(* IEC 61131-3 sources: LASAL/Class/_DriveMngBase (part 2) *)

           ret_code := READY;

           // Daten werden gelöscht :
           L2Buffer[IntRdIndex].AxisNo := 0;
           L2Buffer[IntRdIndex].bActive := FALSE;
           L2NewEntry -= 1;
           if L2NewEntry < 0 then
            L2NewEntry := 0;
           end_if;
           exit;
        end_if;
      end_for;

    end_if;

  else
    ret_code := NewInst(pPara, pResult);
  end_case;

END_FUNCTION

FUNCTION GLOBAL _DriveMngBase::GetAxisWrPtr
	VAR_INPUT
		usAxis 	: USINT;
	END_VAR
	VAR_OUTPUT
		ptr 	: ^_VaranDriveBase::t_WriteValuePtr;
	END_VAR
  VAR
    MyPara   : CmdStruct;
    MyResult : results;
  END_VAR

  if usAxis >= 0 & usAxis < SDDMAXENTRIES then //HasHan
    if bVaranConnected then
      ptr := toVaran.GetAxisWrPtr(AxisNr:=AxBuffer[usAxis].AxisIndex);
    else
      MyPara.uiCmd    := BUSIF_DRIVEMNGBASE_GET_AXIS_WR_PTR;
      MyPara.aPara[0] := to_dint(AxBuffer[usAxis].AxisIndex);
      ToBusIF.NewInst(#MyPara, #MyResult);
      ptr := MyResult.aData[0]$^_VaranDriveBase::t_WriteValuePtr;
    end_if;
  end_if;

END_FUNCTION

FUNCTION GLOBAL _DriveMngBase::GetAxisRdPtr
	VAR_INPUT
		usAxis 	: USINT;
	END_VAR
	VAR_OUTPUT
		ptr 	: ^_VaranDriveBase::t_ReadValuePtr;
	END_VAR
  VAR
    MyPara   : CmdStruct;
    MyResult : results;
  END_VAR

  if usAxis >= 0 & usAxis < SDDMAXENTRIES then //HasHan
    if bVaranConnected then
      ptr := toVaran.GetAxisRdPtr(AxisNr:=AxBuffer[usAxis].AxisIndex);
    else
      MyPara.uiCmd    := BUSIF_DRIVEMNGBASE_GET_AXIS_RD_PTR;
      MyPara.aPara[0] := to_dint(AxBuffer[usAxis].AxisIndex);
      ToBusIF.NewInst(#MyPara, #MyResult);
      ptr := MyResult.aData[0]$^_VaranDriveBase::t_ReadValuePtr;
    end_if;
  end_if;

END_FUNCTION

FUNCTION GLOBAL _DriveMngBase::InitDrive
	VAR_INPUT
		Mode 	: USINT;
	END_VAR
  VAR
    UserPara     : CmdStruct;
    UserResult   : Results;
    x            : USINT;
    pThisNewInst : ^void;
  END_VAR

  if bVaranConnected then
    toVaran.InitDrive();
  else
    UserPara.uiCmd := BUSIF_DRIVEMNGBASE_INIT_DRIVE;
    ToBusIF.NewInst(#UserPara, #UserResult);
  end_if;

  for x := 0 to (SDDMAXENTRIES - 1) do
    if (AxBuffer[x].pThis <> NIL) then
      if (AxBuffer[x].AxisOk = 1) then
        if Mode = 0 then
          UserPara.uiCmd := SDD_INITAXLE;
        else
          UserPara.uiCmd := SDD_URINITAXLE;
        end_if;

        pThisNewInst := AxBuffer[x].pThis;
        pThisNewInst$^VirtualBase^.NewInst(#UserPara, #UserResult);
      end_if;
    end_if;
  end_for;

END_FUNCTION

FUNCTION _DriveMngBase::GetAxIndex
	VAR_INPUT
		AxisNo 	: USINT;
	END_VAR
	VAR_OUTPUT
		AxIndex 	: USINT;
	END_VAR
  VAR
  	x     : USINT;
  END_VAR

  AxIndex := 16#FF;

  for x := 0 to (SDDMAXENTRIES - 1) do
    if (AxBuffer[x].pThis <> NIL) then
      if (AxBuffer[x].AxisOk = 1) & (AxBuffer[x].AxisIndex = AxisNo) then
        AxIndex := x;
        exit;
      end_if;
    else
      exit;
    end_if;
  end_for;

END_FUNCTION

FUNCTION _DriveMngBase::GetAxIndexByAxisBit
	VAR_INPUT
		AxisBit 	: BDINT;
	END_VAR
	VAR_OUTPUT
		AxIndex 	: USINT;
	END_VAR
  VAR
  	x     : USINT;
  END_VAR

  AxIndex := 16#FF;

  for x := 0 to (SDDMAXENTRIES - 1) do
    if (AxBuffer[x].pThis <> NIL) then
      if (AxBuffer[x].AxisBit = AxisBit) then
        AxIndex := x;
        exit;
      end_if;
    else
      exit;
    end_if;
  end_for;

END_FUNCTION

FUNCTION _DriveMngBase::GetFirstAxIndex
	VAR_OUTPUT
		AxIndex 	: USINT;
	END_VAR
  VAR
  	x     : USINT;
  END_VAR

  AxIndex := 16#FF;

  for x := 0 to (SDDMAXENTRIES - 1) do
    if (AxBuffer[x].pThis <> NIL) then
      if (AxBuffer[x].AxisOk = 1) then
        AxIndex := x;
        exit;
      end_if;
    else
      exit;
    end_if;
  end_for;

END_FUNCTION

FUNCTION _DriveMngBase::SetFwVersion
VAR
	szValue     : ARRAY[0..19] of CHAR;
  StrLen      : UDINT;
END_VAR

  Bin2Ascii(pt:=#szValue[0], value:=FwVersionInt, format:=16#820);
  StrLen := _strlen(#szValue[0]);
  FwNumStr.WriteDataOff(udLen:= Strlen, udOff:=0, pData:= #szValue[0]);

END_FUNCTION

FUNCTION _DriveMngBase::SetFwDate
VAR
	szValue     : ARRAY[0..19] of CHAR;
  szFwDate    : ARRAY[0..99] of CHAR;
  StrLen      : UDINT;
  Value       : UDINT;
  tmpYear     : UDINT;
END_VAR

  // Ermitteln des Tages
  Value := FWDateInt AND 16#003F0000;
  Value := Value SHR 16;
  Bin2Ascii(pt:=#szValue[0], value:=Value$DINT, format:=16#102);
  _strcpy(#szFwDate[0], #szValue[0]);
  _strcat(#szFwDate[0], ".");

  // ermitteln des Monats
  Value := FWDateInt AND 16#0F000000;
  Value := Value SHR 24;
  Bin2Ascii(pt:=#szValue[0], value:=Value$DINT, format:=16#102);
  _strcat(#szFwDate[0], #szValue[0]);
  _strcat(#szFwDate[0], ".");

  // ermitteln des Jahres
  Value := FWDateInt AND 16#F0000000;
  Value := Value SHR 28;

  //Newer firmwares >= 2016 are using 2 Bits more, which where originally reserved for day, to have more bits to display year dates.
  //With this change we can display year dates until 2063 instead of 2015,
  tmpYear := FWDateInt AND 16#00C00000;
  tmpYear := tmpYear SHR 18; //Shift Right 18 instead of 22 because these two bits are bit 4 and 5 for the year
  Value := Value OR tmpYear;

  Value += 2000;
  Bin2Ascii(pt:=#szValue[0], value:=Value$DINT, format:=16#800);
  _strcat(#szFwDate[0], #szValue[0]);
  _strcat(#szFwDate[0], " ");

  // ermitteln der Stunde
  Value := FWDateInt AND 16#0000FF00;
  Value := Value SHR 8;
  Bin2Ascii(pt:=#szValue[0], value:=Value$DINT, format:=16#102);
  _strcat(#szFwDate[0], #szValue[0]);
  _strcat(#szFwDate[0], ":");

  // ermitteln der Minuten
  Value := FWDateInt AND 16#000000FF;
  Bin2Ascii(pt:=#szValue[0], value:=Value$DINT, format:=16#102);
  _strcat(#szFwDate[0], #szValue[0]);

  StrLen := _strlen(#szFwDate[0]);
  FwDatetr.WriteDataOff(udLen:= Strlen, udOff:=0, pData:= #szFwDate[0]);

END_FUNCTION

(*
Der String kann folgendermaßen formatiert werden.
xxxx 0000 0000 0000     xxxx = keine Funktion.
     .... .... ****     Anzahl der Dezimalstellen.
     .... **** ....     Position des Dezimalpunkts.
     ...* .... ....     Vornullen (Anzahl der Dezimalstellen).
     ..*. .... ....     Nachkomma Nullen.
     .*.. .... ....     Vorzeichen unmittelbar vor wert (-3 ansonsten - 3).
     *... .... ....     Anzahl der Stellen automatisch ermitteln.

*)

FUNCTION _DriveMngBase::Bin2Ascii
	VAR_INPUT
		pt 	: ^CHAR;
		value 	: DINT;
		format 	: BINT;
	END_VAR
VAR
	tmp		: DINT;
	nk		: UINT;
	dig		: UINT;
	hp     : ^CHAR;
	pd     : UINT;
	h      : UINT;
END_VAR

	if((format AND 16#000F) = 0) then
		format := format OR 16#0800;
	end_if;

	if(format AND 16#0800) then
		tmp  := value;
		if tmp = 0 then
			dig := 1;
		else
			dig := 0;
		end_if;

	    while(tmp) do

			tmp := tmp / 10;
			dig += 1;
	    end_while;

	    nk := ((format SHR 4) AND 16#0F);

		if(nk >= dig) then
	      dig := nk + 1;
		end_if;

		format := (format AND 16#FFF0) OR (dig AND 16#000F);
	end_if;

  dig := (format and 16#0F);		// Anzahl der Stellen
  hp  := pt + dig; 					// pointer auf String-Ende
  tmp := value; 					// Zahl
  pd  := (format shr 4) and 16#0F;	// position des Komma

  if(value < 0) then  		// kontrolle ob Zahl negativ
	hp    += 1;
    value := -value;		// Zahl * (-1)
    pt^   := '-';			// Erstes Zeichen auf '-' setzen
  end_if;

  if(format and 16#0200) then   // Nachnullen löschen
    h := pd;
	while(h) do					// Nur Nullen hinter Komma
	  h -= 1;
	  if((value mod 10) = 0) then	// Ist Ziffer Null?
	    value := value / 10; 	// wenn ja, Null löschen
		pd -= 1;
      else
	    h := 0;
      end_if;

	end_while;
  end_if;

  if(pd <> 0) then    	// Komma noch zu setzen?
    hp += 1;
  end_if;

  hp^ := 0;           	// String mit Ascii-0 abschließen
  hp  -= 1;

  repeat
    hp^   := '0' + TO_USINT(value mod 10); //akt. Ziffer
	hp    -= 1;
	pd    -= 1;
	dig   -= 1;
	if(pd = 0)then		//	Komma setzen?
	  hp^ := '.';
	  hp -= 1;
    end_if;

    value := value / 10; 	// nächste Ziffer

    if((dig = 0) & (value <> 0)) then	// Zahl zu groß
	  pt^   := '?'; 	// Formatfehler
	  value := 0;
	end_if;
  until(value = 0) end_repeat;

  if(dig > 0) then 	// mit Vornullen auffüllen
	repeat			// so lange bis Digits auf Null
      if((format and 16#0100)|(pd$INT >= 0)) then   // Vornullen im
        hp^ := '0'; 								// Format angegeben?
      else			// formatfehler (digit zu groß und keine Vornullen)
	    pt^   := '?'; 	// Formatfehler
	    value := 0;
      end_if;
      pd -= 1;
	  hp -= 1;
      if(pd = 0) then	// Komma setzen
	    hp^ := '.';
	    hp -= 1;
      end_if;
	  dig -= 1;
	until(dig = 0) end_repeat; 	// letzte Ziffer?
  end_if;

END_FUNCTION

FUNCTION VIRTUAL GLOBAL _DriveMngBase::RetryCounter::Read
	VAR_OUTPUT
		output (EAX) 	: UDINT;
	END_VAR
  VAR
    MyPara   : CmdStruct;
    MyResult : results;
  END_VAR

  if bVaranConnected then
    RetryCounter := toVaran.RetryCounter.Read();
  else
    MyPara.uiCmd  := BUSIF_DRIVEMNGBASE_READ_RETRY_COUNTER;
    ToBusIF.NewInst(#MyPara, #MyResult);
    RetryCounter := MyResult.aData[0]$UDINT;
  end_if;

  output := RetryCounter;

END_FUNCTION

FUNCTION GLOBAL _DriveMngBase::SetSyncEntry
	VAR_INPUT
		usAxis 	: USINT;
		usValue 	: USINT;
		usPData 	: DINT;
	END_VAR
	VAR_OUTPUT
		retcode 	: DINT;
	END_VAR
  VAR
    MyPara   : CmdStruct;
    MyResult : results;
  END_VAR

  if usAxis >= 0 & usAxis < SDDMAXENTRIES then //HasHan
    if bVaranConnected then
      retcode:=toVaran.SetSyncParameter(us_Axis:=AxBuffer[usAxis].AxisIndex, us_value:=usValue, sd_data:=usPData);
    else
      MyPara.uiCmd    := BUSIF_DRIVEMNGBASE_SET_SYNC_PARA;
      MyPara.aPara[0] := to_dint(AxBuffer[usAxis].AxisIndex);
      MyPara.aPara[1] := to_dint(usValue);
      MyPara.aPara[2] := to_dint(usPData);

      ToBusIF.NewInst(#MyPara, #MyResult);
      retcode := MyResult.aData[0]$DINT;
    end_if;
  else
    retcode := -1;
  end_if;

END_FUNCTION

FUNCTION GLOBAL _DriveMngBase::GetSyncEntry
	VAR_INPUT
		usAxis 	: USINT;
		usValue : USINT;
		usPData : ^DINT;
	END_VAR
	VAR_OUTPUT
		retcode : DINT;
	END_VAR
  VAR
    MyPara   : CmdStruct;
    MyResult : results;
  END_VAR

  if usAxis >= 0 & usAxis < SDDMAXENTRIES then //HasHan
    if bVaranConnected then
      retcode:=toVaran.GetSyncParameter(us_Axis:=AxBuffer[usAxis].AxisIndex, us_value:=usValue, p_data:=usPData);
    else
      MyPara.uiCmd    := BUSIF_DRIVEMNGBASE_GET_SYNC_PARA;
      MyPara.aPara[0] := to_dint(AxBuffer[usAxis].AxisIndex);
      MyPara.aPara[1] := to_dint(usValue);
      MyPara.aPara[2] := (usPData)$DINT;

      ToBusIF.NewInst(#MyPara, #MyResult);
      retcode := MyResult.aData[0]$DINT;
    end_if;
  else
    retcode := -1;
  end_if;

END_FUNCTION

FUNCTION _DriveMngBase::GetDriveType
	VAR_INPUT
		HWCode 	: DINT;
	END_VAR
	VAR_OUTPUT
		DriveType 	: _DRIVETYPE;
	END_VAR
  VAR
  	buffer   : DINT;
    MyPara   : CmdStruct;
    MyResult : results;
    dRetCode : iprStates;
  END_VAR

  if bVaranConnected then
    buffer := HWCode SHR 16;
    case buffer of
    // 3 Achsen
      0: DriveType:=_SDD_310;
      1: DriveType:=_SDD_315;
      2: DriveType:=_S_340;
      3: DriveType:=_SDD_310;
      4: DriveType:=_S_340;
      6: DriveType:=_SDD_315;
     12: DriveType:=_SDD_335;
     16: DriveType:=_SDD_305;
     20: DriveType:=_SDD_305;
     26: DriveType:=_SDD_310;

     // 2 Achsen
      5: DriveType:=_SDD_215;
      9: DriveType:=_SDD_210;
     22: DriveType:=_SDD_205;

     // 1 Achse
      7: DriveType:=_SDD_120;
     21: DriveType:=_SDD_105;
     10: DriveType:=_SDD_115;

    else
      DriveType:=_NotFound;
    end_case;

  else
    //if businterface is connected
    MyPara.uiCmd    := BUSIF_DRIVEMNGBASE_GET_BUSTYPE;
    //first parameter is the length of followed data
    MyPara.aPara[0] := 0;

    dRetCode := ToBusIF.NewInst(#MyPara, #MyResult);

    if dRetCode = Ready
    & MyResult.uiLng = 1 then
      if MyResult.aData[0] = HWT_ESCAPE_SDIAS then
        case DeviceID of
          DRIVEMNG_BUSDEVICEID_DC061:
            DriveType := _DC061;

          DRIVEMNG_BUSDEVICEID_DC062:
            DriveType := _DC062;

        else
          DriveType:=_NotFound;
        end_case;

      elsif MyResult.aData[0] = HWT_ESCAPE_VARAN then
        case DeviceID of
          DRIVEMNG_BUSDEVICEID_SDD1300:
            DriveType := _SDD_1300;

          DRIVEMNG_BUSDEVICEID_SDD1400:
            DriveType := _SDD_1400;

          DRIVEMNG_BUSDEVICEID_SDD1500:
            DriveType := _SDD_1500;

          DRIVEMNG_BUSDEVICEID_SDD1600:
            DriveType := _SDD_1600;

        else
          DriveType:=_NotFound;

        end_case;

      elsif MyResult.aData[0] = HWT_ESCAPE_VARAN_S2 then
        case DeviceID of

          DRIVEMNG_BUSDEVICEID_WA011:
            DriveType := _WA011;

          DRIVEMNG_BUSDEVICEID_WA012:
            DriveType := _WA012;

        else
          DriveType:=_NotFound;

        end_case;

      else
        DriveType:=_NotFound;
      end_if;

    else
      DriveType:=_NotFound;
    end_if;
  end_if;

END_FUNCTION

FUNCTION GLOBAL _DriveMngBase::GetVaranDriveState
	VAR_OUTPUT
		retcode 	: DINT;
	END_VAR
  VAR
    MyPara   : CmdStruct;
    MyResult : results;
  END_VAR

  if bVaranConnected then
    retcode := toVaran.GetDriveIntState();
  else
    MyPara.uiCmd := BUSIF_DRIVEMNGBASE_GET_DRIVE_INT_STATE;
    ToBusIF.NewInst(#MyPara, #MyResult);
    retcode := MyResult.aData[0]$DINT;
  end_if;

END_FUNCTION

FUNCTION GLOBAL _DriveMngBase::SetTimeBase
	VAR_INPUT
		ud_timebase_ms 	: UDINT;
	END_VAR
	VAR_OUTPUT
		sd_retval 	: DINT;
	END_VAR

  //When the DriveMng is called manuelly instead of setting the CyWork Time,
  //the Customer has to tell the Class, witch TimeBase is set, because this Time is use somewhere in the Class.

  IF InitCounter <= 1 THEN  //The Init use the ud_TimeoutCycles and set any value, to prevent
                            //the override from this Value after the Customer has set the TimeBase manuelly, this Methode only works after the first Init run.
    sd_retval := -1;
  else
    IF ud_timebase_ms <> 0 THEN
      ud_timebase_ms *= 1000; // Rev. 1.16: us is the unit for the calculation
      ud_TimeoutCycles := ( SDD_ASY_TIMEOUT / ud_timebase_ms ) + 5;
      sd_retval := 0;
    ELSE
      sd_retval := -2;
    END_IF;
  END_IF;

END_FUNCTION

FUNCTION _DriveMngBase::_DriveMngBase
	VAR_OUTPUT
		ret_code 	: ConfStates;
	END_VAR

  //Rev. 1.16: to avoid wrong information on server if drive is used as a transparent client
  CmdState := _NotInitialized;

	ret_code := C_OK;

END_FUNCTION

FUNCTION VIRTUAL _DriveMngBase::GetBusDeviceID
	VAR_OUTPUT
		output 	: UDINT;
	END_VAR

  //Overwrite this method in derived class
  output := HWC_INVALID_DEVICE_ID;

END_FUNCTION

FUNCTION VIRTUAL _DriveMngBase::GetDrvDeviceID
	VAR_OUTPUT
		output 	: UDINT;
	END_VAR

  //Overwrite this method in derived class
  output := HWC_INVALID_DEVICE_ID;

END_FUNCTION

FUNCTION GLOBAL _DriveMngBase::IsAnyAxisEnabled
	VAR_OUTPUT
		AnyAxisEnabled 	: BOOL;
	END_VAR
  VAR
    UserPara     : CmdStruct;
    UserResult   : Results;
    x            : USINT;
    pThisNewInst : ^void;
  END_VAR

  // search for any enabled axis (all axis must be disabled to set absolut position, because drive needs to switch communication)
  AnyAxisEnabled := FALSE;
  UserPara.uiCmd := SDD_GET_ANY_AXIS_ENABLED;

  for x := 0 to (SDDMAXENTRIES - 1) do
    if (AxBuffer[x].pThis <> NIL) then
      if (AxBuffer[x].AxisOk = 1) then
        UserResult.uiLng := 0;

        pThisNewInst := AxBuffer[x].pThis;
        pThisNewInst$^VirtualBase^.NewInst(#UserPara, #UserResult);

        // if there is an enabled axis
        if (UserResult.uiLng = 1) & UserResult.aData[0] then
          // leave method
          AnyAxisEnabled := TRUE;
          return;
        end_if;
      end_if;
    end_if;
  end_for;

END_FUNCTION

FUNCTION GLOBAL _DriveMngBase::DisableDevice
	VAR_OUTPUT
		RetCode 	: DINT;
	END_VAR
  VAR
    MyPara   : CmdStruct;
    MyResult : results;
  END_VAR

  if bVaranConnected then
    RetCode := toVaran.DisableDevice();
  else
    MyPara.uiCmd    := BUSIF_DRIVEMNGBASE_WRITE_PARAMETER;
    Mypara.aPara[0] := _BUS_IF_DRVMNG_DISABLE_DEVICE;
    RetCode$UDINT   := ToBusIF.NewInst(#MyPara, #MyResult);
    if RetCode$IprStates = ERROR then
      RetCode := -1;
    end_if;
  end_if;

END_FUNCTION

FUNCTION GLOBAL _DriveMngBase::EnableDevice
	VAR_OUTPUT
		RetCode 	: DINT;
	END_VAR
  VAR
    MyPara   : CmdStruct;
    MyResult : results;
  END_VAR

  if bVaranConnected then
    RetCode := toVaran.EnableDevice();
  else
    MyPara.uiCmd    := BUSIF_DRIVEMNGBASE_WRITE_PARAMETER;
    Mypara.aPara[0] := _BUS_IF_DRVMNG_ENABLE_DEVICE;
    RetCode$UDINT   := ToBusIF.NewInst(#MyPara, #MyResult);
    if RetCode$IprStates = ERROR then
      RetCode := -1;
    end_if;
  end_if;

END_FUNCTION
